REGION Network 1: Header
   // ==============================================================================
   //  Company: Precision Automation & Robotics India Ltd. 
   // ------------------------------------------------------------------------------
   //  Item Code: S21006022015
   //  Author/Created by: Manoj Sonawane
   //  Reviewed/Checked by: Sandip.c
   //  First Release on: 19-07-24
   //  Latest update on:11-03-25
   // ------------------------------------------------------------------------------
   //  Tested with: CPU firmware, model or simulator testing
   //  Engineering/Editor: TIA Portal V17
   // ------------------------------------------------------------------------------
   //  Restrictions:
   //  Dependencies/Requirements:
   //  1. "UDT_IS28xx_To_Plc"
   //  2. "UDT_Plc_To_IS28xx"
   // ------------------------------------------------------------------------------
   //  Change Log:
   //  Ver.	Date		Changed by		Details of changes
   //  1.0	 19-07-24                 Manoj Sonawane            	First release version
   // 1.1              30-09-24                 Harshal Gharmode                         Modify as per shop floor testing
   // 1.2              11-03-25                 Swapnil Asule                                  Remove retry count logic & update                                                                                                                         data Inspection logic
   // ------------------------------------------------------------------------------
   //  Functionality:  : The Cognex In-Sight® 2801 vision system communicates with the Siemence s7-15xx series PLC over Profinet protocol.The main functionality of this block is provided for the user can change the job ID according to their needs and get the inspection result data of Job ID.
   // 
   // 
   //  Inputs
   // iInsightCamera_Input	"UDT_IS28xx_To_Plc"
   // iResetFault	Bool
   // iModuleReset	Bool
   // iAutorunning	Bool
   // iStartJobSelection	Bool
   // iStartInspection	Bool
   // iJobID	Int
   // iUserData	Array[1..60] of Byte
   // iTriggerEnableTimeoutTime	Time
   // iTriggerTimeoutTime	Time
   // iAcquiringTimeOutTime	Time
   // iPrgmNoTimeOut	Time
   // iFeedbackTimeOut	Time
   // 
   //  Outputs
   //  qInsightCamera_Output	"UDT_Plc_To_IS28xx"
   // qJobPass	Bool
   // qJobFail	Bool
   // qJobSelectionOver	Bool
   // qJobInspectionOver	Bool
   // qVisionOnline	Bool
   // qVisionOfflineReason1	Bool
   // qVisionOfflineReason2	Bool
   // qVisionOfflineReason3	Bool
   // qErrBothStartOn	Bool
   // qErrJobSelection	Bool
   // qErrTriggerEnableTimeout	Bool
   // qErrTriggerTimeOut	Bool
   // qErrAcquiringTimeOut	Bool
   // qErrJobIDEchoMismatch	Bool
   // qErrSetUserDataAckNtRcvd	Bool
   // qMsgJobIDMismatch	Bool
   // qInspectionResult	Array[1..60] of Byte
   // 
   //  In-outs
   //  iqRunningJobID	Int
   // ------------------------------------------------------------------------------
   //  Errors reported:
   //  1.qErrTriggerTimeO : Error trigger timeout
   //  2. qErrAcquiringTimeOut;Acquiring Time Out
   //  3. qErrTriggerEnableTimeout:Trigger Enable Time Out
   //  4. qErrJobSelection: Job selection error
   //  5. qErrBothStartOn: Start Inspection & Start Job Selection command are active at same time
   //  6. qErrJobIDEchoMismatch: Set Job ID & its echo is not matched
   //  7. qErrSetUserDataAckNtRcvd: Set user data acknowldge not recived within the defined time.
   // 
   //  Messages reported:
   //   1. qMsgJobIDMismatch: Set Job ID & running JOB ID is not matched
   // ==============================================================================
END_REGION

REGION Network 2: Reset Faults
   // Reset Faults
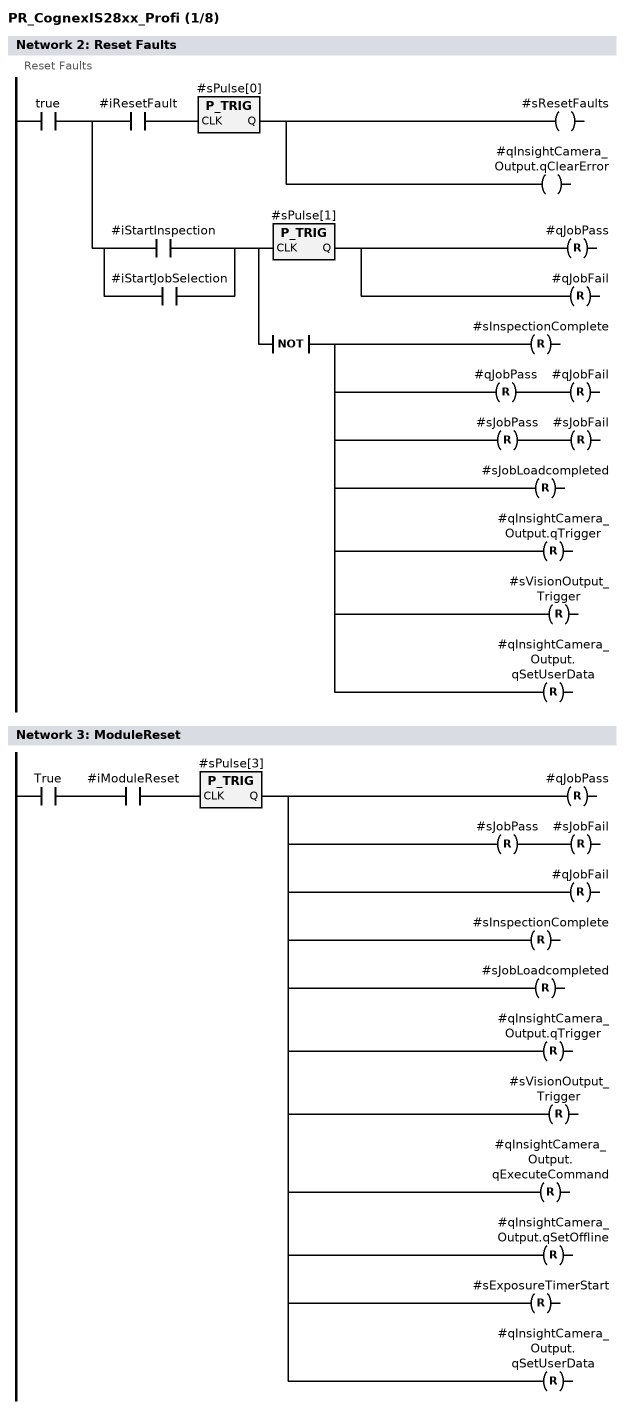
   RUNG wire#powerrail
      Contact( true )
      wire#w1
      Contact( #iResetFault )
      P_Trig( #sPulse[0] )
      wire#w2
      Coil( #sResetFaults )
   END_RUNG
   RUNG wire#w2
      Coil( #qInsightCamera_Output.qClearError )
   END_RUNG
   RUNG wire#w1
      Contact( #iStartInspection )
      wire#w3
      P_Trig( #sPulse[1] )
      wire#w4
      R_Coil( #qJobPass )
   END_RUNG
   RUNG wire#w1
      Contact( #iStartJobSelection )
   END_RUNG wire#w3
   RUNG wire#w4
      R_Coil( #qJobFail )
   END_RUNG
   RUNG wire#w3
      Not()
      wire#w5
      R_Coil( #sInspectionComplete )
   END_RUNG
   RUNG wire#w5
      R_Coil( #qJobPass )
      R_Coil( #qJobFail )
   END_RUNG
   RUNG wire#w5
      R_Coil( #sJobPass )
      R_Coil( #sJobFail )
   END_RUNG
   RUNG wire#w5
      R_Coil( #sJobLoadcompleted )
   END_RUNG
   RUNG wire#w5
      R_Coil( #qInsightCamera_Output.qTrigger )
   END_RUNG
   RUNG wire#w5
      R_Coil( #sVisionOutput_Trigger )
   END_RUNG
   RUNG wire#w5
      R_Coil( #qInsightCamera_Output.qSetUserData )
   END_RUNG
   // the same network as SCL:
   #_w1 := true AND #iResetFault;
   #_w2 := #_w1 AND NOT #sPulse[0];   // rising edge
   #sPulse[0] := #_w1;
   #sResetFaults := #_w2;
   #qInsightCamera_Output.qClearError := #_w2;
   #_w3 := true AND (#iStartInspection OR #iStartJobSelection);
   #_w4 := #_w3 AND NOT #sPulse[1];   // rising edge
   #sPulse[1] := #_w3;
   IF #_w4 THEN
       #qJobPass := FALSE;
       #qJobFail := FALSE;
   END_IF;
   IF NOT #_w3 THEN
       #sInspectionComplete := FALSE;
       #qJobPass := FALSE;
       #qJobFail := FALSE;
       #sJobPass := FALSE;
       #sJobFail := FALSE;
       #sJobLoadcompleted := FALSE;
       #qInsightCamera_Output.qTrigger := FALSE;
       #sVisionOutput_Trigger := FALSE;
       #qInsightCamera_Output.qSetUserData := FALSE;
   END_IF;
END_REGION

REGION Network 3: ModuleReset
   RUNG wire#powerrail
      Contact( True )
      Contact( #iModuleReset )
      P_Trig( #sPulse[3] )
      wire#w1
      R_Coil( #qJobPass )
   END_RUNG
   RUNG wire#w1
      R_Coil( #sJobPass )
      R_Coil( #sJobFail )
   END_RUNG
   RUNG wire#w1
      R_Coil( #qJobFail )
   END_RUNG
   RUNG wire#w1
      R_Coil( #sInspectionComplete )
   END_RUNG
   RUNG wire#w1
      R_Coil( #sJobLoadcompleted )
   END_RUNG
   RUNG wire#w1
      R_Coil( #qInsightCamera_Output.qTrigger )
   END_RUNG
   RUNG wire#w1
      R_Coil( #sVisionOutput_Trigger )
   END_RUNG
   RUNG wire#w1
      R_Coil( #qInsightCamera_Output.qExecuteCommand )
   END_RUNG
   RUNG wire#w1
      R_Coil( #qInsightCamera_Output.qSetOffline )
   END_RUNG
   RUNG wire#w1
      R_Coil( #sExposureTimerStart )
   END_RUNG
   RUNG wire#w1
      R_Coil( #qInsightCamera_Output.qSetUserData )
   END_RUNG
   // the same network as SCL:
   #_w1 := True AND #iModuleReset;
   #_w2 := #_w1 AND NOT #sPulse[3];   // rising edge
   #sPulse[3] := #_w1;
   IF #_w2 THEN
       #qJobPass := FALSE;
       #sJobPass := FALSE;
       #sJobFail := FALSE;
       #qJobFail := FALSE;
       #sInspectionComplete := FALSE;
       #sJobLoadcompleted := FALSE;
       #qInsightCamera_Output.qTrigger := FALSE;
       #sVisionOutput_Trigger := FALSE;
       #qInsightCamera_Output.qExecuteCommand := FALSE;
       #qInsightCamera_Output.qSetOffline := FALSE;
       #sExposureTimerStart := FALSE;
       #qInsightCamera_Output.qSetUserData := FALSE;
   END_IF;
END_REGION

REGION Network 4: Time out validation
   // Time out validation 1. Trigger enable time out
   // 2. Trigger time out
   // 3. Acquiring TimeOut Time
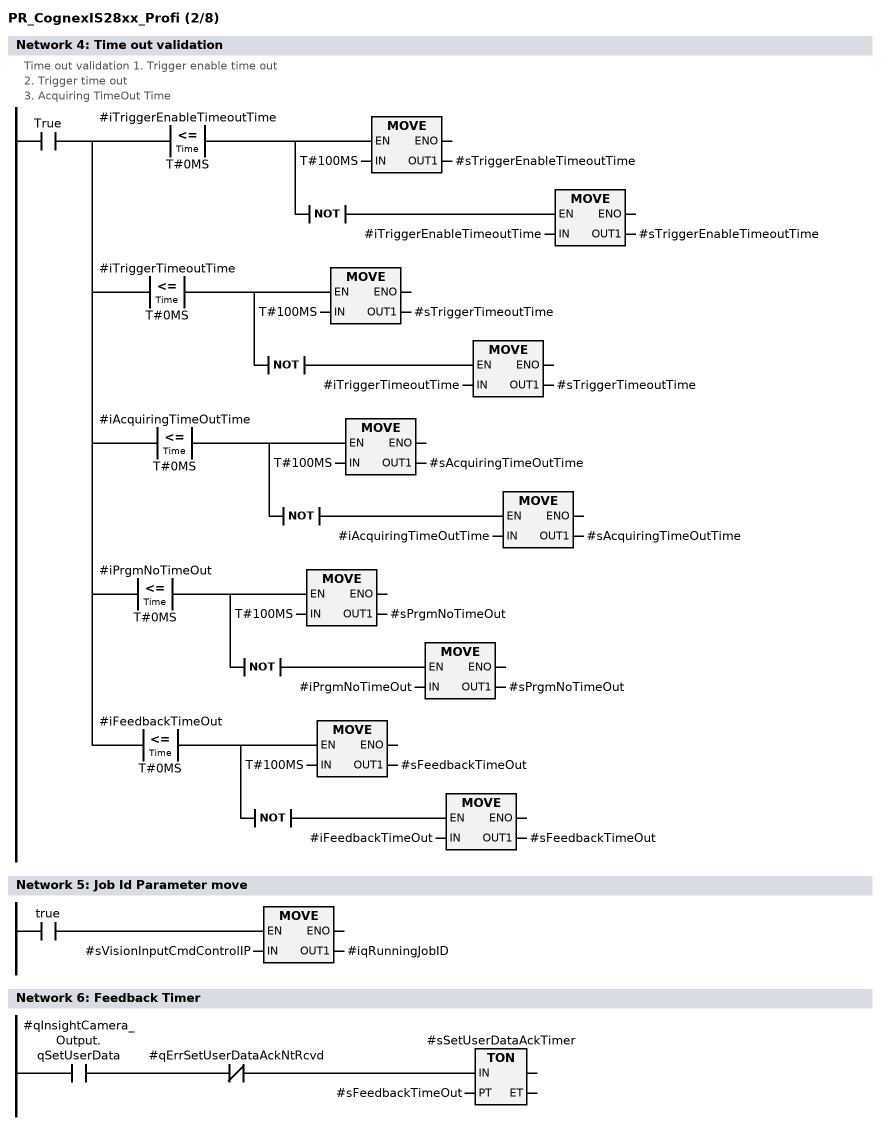
   RUNG wire#powerrail
      Contact( True )
      wire#w1
      { S7_Templates := "SrcType := Time" } LE_Contact(in1 := #iTriggerEnableTimeoutTime, in2 := T#0MS)
      wire#w2
      Move(in := T#100MS, out1 => #sTriggerEnableTimeoutTime)
   END_RUNG
   RUNG wire#w2
      Not()
      Move(in := #iTriggerEnableTimeoutTime, out1 => #sTriggerEnableTimeoutTime)
   END_RUNG
   RUNG wire#w1
      { S7_Templates := "SrcType := Time" } LE_Contact(in1 := #iTriggerTimeoutTime, in2 := T#0MS)
      wire#w3
      Move(in := T#100MS, out1 => #sTriggerTimeoutTime)
   END_RUNG
   RUNG wire#w3
      Not()
      Move(in := #iTriggerTimeoutTime, out1 => #sTriggerTimeoutTime)
   END_RUNG
   RUNG wire#w1
      { S7_Templates := "SrcType := Time" } LE_Contact(in1 := #iAcquiringTimeOutTime, in2 := T#0MS)
      wire#w4
      Move(in := T#100MS, out1 => #sAcquiringTimeOutTime)
   END_RUNG
   RUNG wire#w4
      Not()
      Move(in := #iAcquiringTimeOutTime, out1 => #sAcquiringTimeOutTime)
   END_RUNG
   RUNG wire#w1
      { S7_Templates := "SrcType := Time" } LE_Contact(in1 := #iPrgmNoTimeOut, in2 := T#0MS)
      wire#w5
      Move(in := T#100MS, out1 => #sPrgmNoTimeOut)
   END_RUNG
   RUNG wire#w5
      Not()
      Move(in := #iPrgmNoTimeOut, out1 => #sPrgmNoTimeOut)
   END_RUNG
   RUNG wire#w1
      { S7_Templates := "SrcType := Time" } LE_Contact(in1 := #iFeedbackTimeOut, in2 := T#0MS)
      wire#w6
      Move(in := T#100MS, out1 => #sFeedbackTimeOut)
   END_RUNG
   RUNG wire#w6
      Not()
      Move(in := #iFeedbackTimeOut, out1 => #sFeedbackTimeOut)
   END_RUNG
   // the same network as SCL:
   #_w1 := True AND (#iTriggerEnableTimeoutTime <= T#0MS);
   IF #_w1 THEN #sTriggerEnableTimeoutTime := T#100MS; END_IF;
   IF NOT #_w1 THEN #sTriggerEnableTimeoutTime := #iTriggerEnableTimeoutTime; END_IF;
   #_w2 := True AND (#iTriggerTimeoutTime <= T#0MS);
   IF #_w2 THEN #sTriggerTimeoutTime := T#100MS; END_IF;
   IF NOT #_w2 THEN #sTriggerTimeoutTime := #iTriggerTimeoutTime; END_IF;
   #_w3 := True AND (#iAcquiringTimeOutTime <= T#0MS);
   IF #_w3 THEN #sAcquiringTimeOutTime := T#100MS; END_IF;
   IF NOT #_w3 THEN #sAcquiringTimeOutTime := #iAcquiringTimeOutTime; END_IF;
   #_w4 := True AND (#iPrgmNoTimeOut <= T#0MS);
   IF #_w4 THEN #sPrgmNoTimeOut := T#100MS; END_IF;
   IF NOT #_w4 THEN #sPrgmNoTimeOut := #iPrgmNoTimeOut; END_IF;
   #_w5 := True AND (#iFeedbackTimeOut <= T#0MS);
   IF #_w5 THEN #sFeedbackTimeOut := T#100MS; END_IF;
   IF NOT #_w5 THEN #sFeedbackTimeOut := #iFeedbackTimeOut; END_IF;
END_REGION

REGION Network 5: Job Id Parameter move
   RUNG wire#powerrail
      Contact( true )
      Move(in := #sVisionInputCmdControlIP, out1 => #iqRunningJobID)
   END_RUNG
   // the same network as SCL:
   IF true THEN #iqRunningJobID := #sVisionInputCmdControlIP; END_IF;
END_REGION

REGION Network 6: Feedback Timer
   #sSetUserDataAckTimer(IN := #qInsightCamera_Output.qSetUserData AND NOT #qErrSetUserDataAckNtRcvd,   // TON
                         PT := #sFeedbackTimeOut);
END_REGION

REGION Network 7: UserData
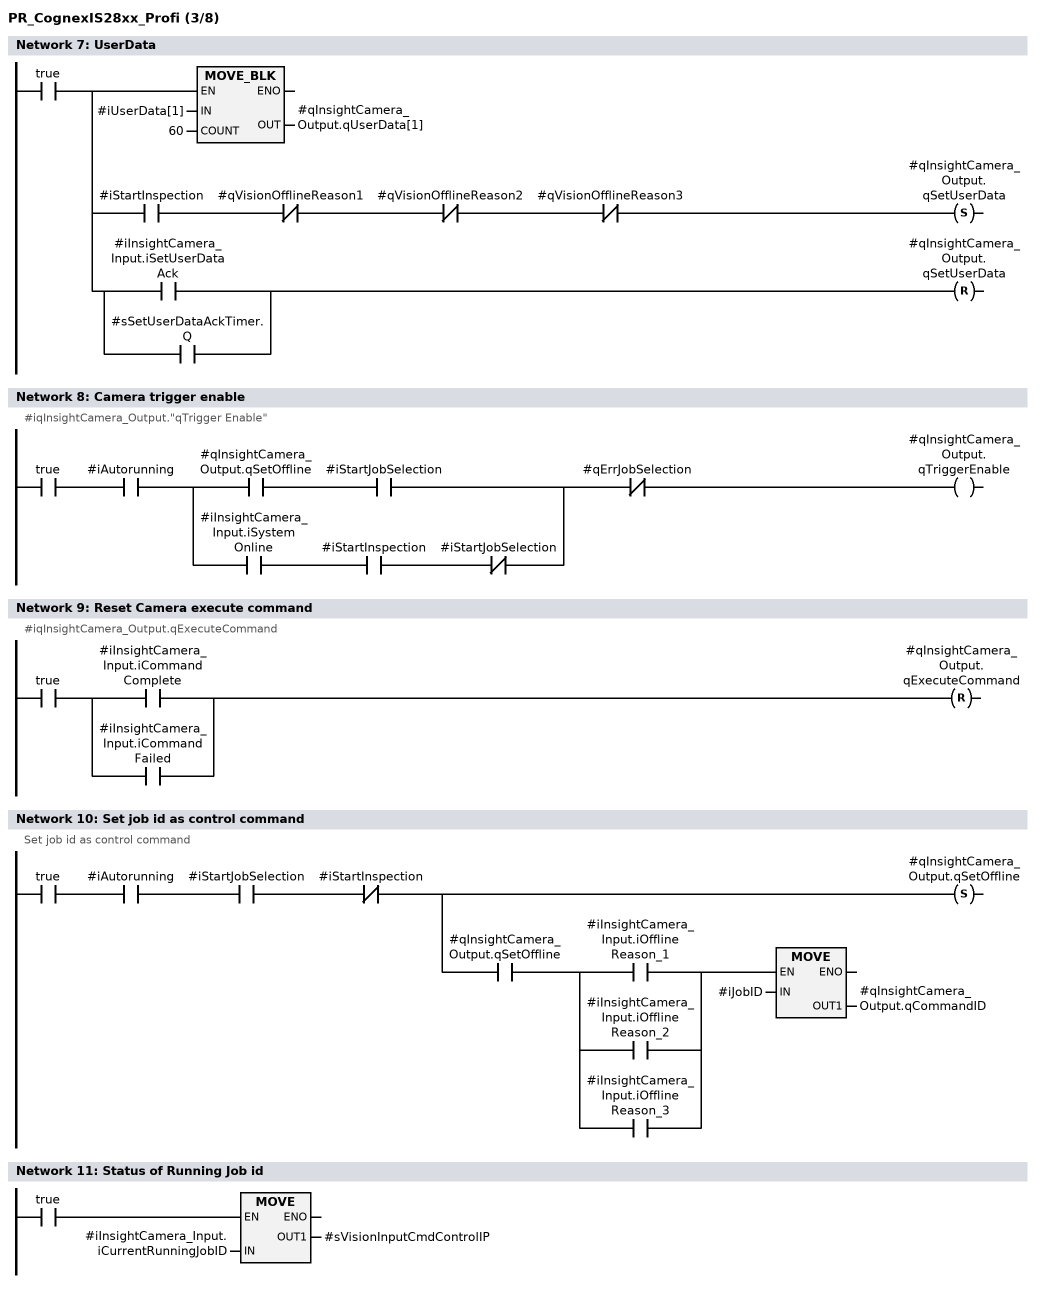
   IF true THEN
       MOVE_BLK(IN := #iUserData[1], COUNT := 60, OUT => #qInsightCamera_Output.qUserData[1]);
   END_IF;
   IF true AND #iStartInspection AND NOT #qVisionOfflineReason1 AND NOT #qVisionOfflineReason2 AND NOT #qVisionOfflineReason3 THEN
       #qInsightCamera_Output.qSetUserData := TRUE;
   END_IF;
   IF true AND (#iInsightCamera_Input.iSetUserDataAck OR #sSetUserDataAckTimer.Q) THEN
       #qInsightCamera_Output.qSetUserData := FALSE;
   END_IF;
END_REGION

REGION Network 8: Camera trigger enable
   // #iqInsightCamera_Output."qTrigger Enable"
   RUNG wire#powerrail
      Contact( true )
      Contact( #iAutorunning )
      wire#w1
      Contact( #qInsightCamera_Output.qSetOffline )
      Contact( #iStartJobSelection )
      wire#w2
      I_Contact( #qErrJobSelection )
      Coil( #qInsightCamera_Output.qTriggerEnable )
   END_RUNG
   RUNG wire#w1
      Contact( #iInsightCamera_Input.iSystemOnline )
      Contact( #iStartInspection )
      I_Contact( #iStartJobSelection )
   END_RUNG wire#w2
   // the same network as SCL:
   #qInsightCamera_Output.qTriggerEnable := true AND #iAutorunning AND ((#qInsightCamera_Output.qSetOffline AND #iStartJobSelection) OR (#iInsightCamera_Input.iSystemOnline AND #iStartInspection AND NOT #iStartJobSelection)) AND NOT #qErrJobSelection;
END_REGION

REGION Network 9: Reset Camera execute command
   // #iqInsightCamera_Output.qExecuteCommand
   RUNG wire#powerrail
      Contact( true )
      wire#w1
      Contact( #iInsightCamera_Input.iCommandComplete )
      wire#w2
      R_Coil( #qInsightCamera_Output.qExecuteCommand )
   END_RUNG
   RUNG wire#w1
      Contact( #iInsightCamera_Input.iCommandFailed )
   END_RUNG wire#w2
   // the same network as SCL:
   IF true AND (#iInsightCamera_Input.iCommandComplete OR #iInsightCamera_Input.iCommandFailed) THEN
       #qInsightCamera_Output.qExecuteCommand := FALSE;
   END_IF;
END_REGION

REGION Network 10: Set job id as control command
   // Set job id as control command
   RUNG wire#powerrail
      Contact( true )
      Contact( #iAutorunning )
      Contact( #iStartJobSelection )
      I_Contact( #iStartInspection )
      wire#w1
      S_Coil( #qInsightCamera_Output.qSetOffline )
   END_RUNG
   RUNG wire#w1
      Contact( #qInsightCamera_Output.qSetOffline )
      wire#w2
      Contact( #iInsightCamera_Input.iOfflineReason_1 )
      wire#w3
      Move(in := #iJobID, out1 => #qInsightCamera_Output.qCommandID)
   END_RUNG
   RUNG wire#w2
      Contact( #iInsightCamera_Input.iOfflineReason_2 )
   END_RUNG wire#w3
   RUNG wire#w2
      Contact( #iInsightCamera_Input.iOfflineReason_3 )
   END_RUNG wire#w3
   // the same network as SCL:
   #_w1 := true AND #iAutorunning AND #iStartJobSelection AND NOT #iStartInspection;
   IF #_w1 THEN #qInsightCamera_Output.qSetOffline := TRUE; END_IF;
   IF #_w1 AND #qInsightCamera_Output.qSetOffline AND (#iInsightCamera_Input.iOfflineReason_1 OR #iInsightCamera_Input.iOfflineReason_2 OR #iInsightCamera_Input.iOfflineReason_3) THEN
       #qInsightCamera_Output.qCommandID := #iJobID;
   END_IF;
END_REGION

REGION Network 11: Status of Running Job id
   RUNG wire#powerrail
      Contact( true )
      Move(in := #iInsightCamera_Input.iCurrentRunningJobID, out1 => #sVisionInputCmdControlIP)
   END_RUNG
   // the same network as SCL:
   IF true THEN #sVisionInputCmdControlIP := #iInsightCamera_Input.iCurrentRunningJobID; END_IF;
END_REGION

REGION Network 12: Set Execute command as per Job selection
   // Set Execute command as per Job selection
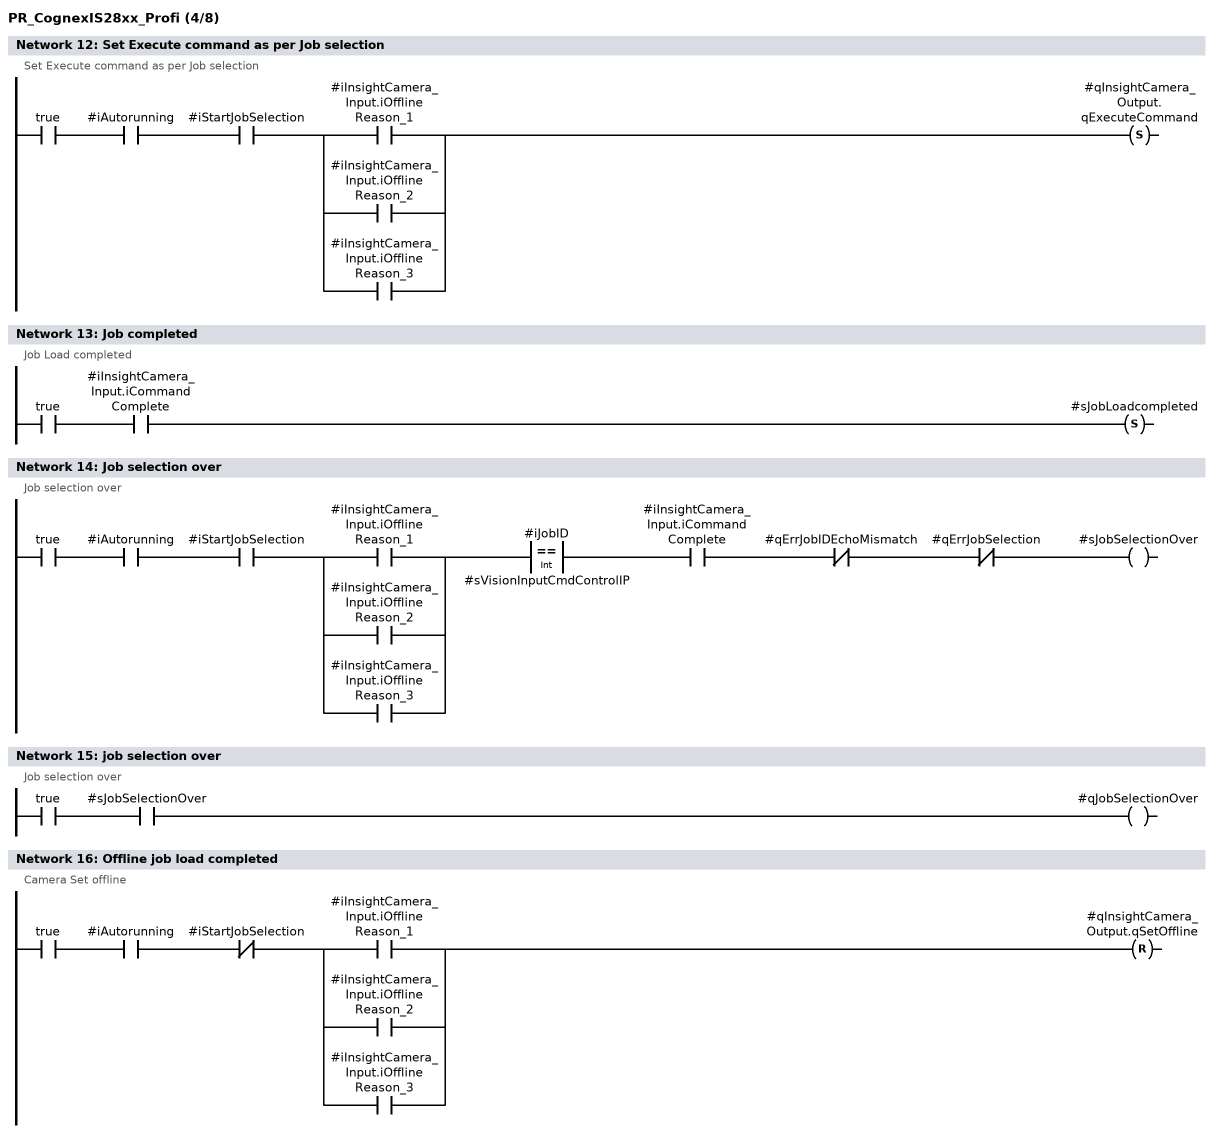
   RUNG wire#powerrail
      Contact( true )
      Contact( #iAutorunning )
      Contact( #iStartJobSelection )
      wire#w1
      Contact( #iInsightCamera_Input.iOfflineReason_1 )
      wire#w2
      S_Coil( #qInsightCamera_Output.qExecuteCommand )
   END_RUNG
   RUNG wire#w1
      Contact( #iInsightCamera_Input.iOfflineReason_2 )
   END_RUNG wire#w2
   RUNG wire#w1
      Contact( #iInsightCamera_Input.iOfflineReason_3 )
   END_RUNG wire#w2
   // the same network as SCL:
   IF true AND #iAutorunning AND #iStartJobSelection AND (#iInsightCamera_Input.iOfflineReason_1 OR #iInsightCamera_Input.iOfflineReason_2 OR #iInsightCamera_Input.iOfflineReason_3) THEN
       #qInsightCamera_Output.qExecuteCommand := TRUE;
   END_IF;
END_REGION

REGION Network 13: Job completed
   // Job Load completed
   RUNG wire#powerrail
      Contact( true )
      Contact( #iInsightCamera_Input.iCommandComplete )
      S_Coil( #sJobLoadcompleted )
   END_RUNG
   // the same network as SCL:
   IF true AND #iInsightCamera_Input.iCommandComplete THEN #sJobLoadcompleted := TRUE; END_IF;
END_REGION

REGION Network 14: Job selection over
   // Job selection over
   RUNG wire#powerrail
      Contact( true )
      Contact( #iAutorunning )
      Contact( #iStartJobSelection )
      wire#w1
      Contact( #iInsightCamera_Input.iOfflineReason_1 )
      wire#w2
      { S7_Templates := "SrcType := Int" } EQ_Contact(in1 := #iJobID, in2 := #sVisionInputCmdControlIP)
      Contact( #iInsightCamera_Input.iCommandComplete )
      I_Contact( #qErrJobIDEchoMismatch )
      I_Contact( #qErrJobSelection )
      Coil( #sJobSelectionOver )
   END_RUNG
   RUNG wire#w1
      Contact( #iInsightCamera_Input.iOfflineReason_2 )
   END_RUNG wire#w2
   RUNG wire#w1
      Contact( #iInsightCamera_Input.iOfflineReason_3 )
   END_RUNG wire#w2
   // the same network as SCL:
   #sJobSelectionOver := true AND #iAutorunning AND #iStartJobSelection AND (#iInsightCamera_Input.iOfflineReason_1 OR #iInsightCamera_Input.iOfflineReason_2 OR #iInsightCamera_Input.iOfflineReason_3) AND (#iJobID = #sVisionInputCmdControlIP) AND #iInsightCamera_Input.iCommandComplete AND NOT #qErrJobIDEchoMismatch AND NOT #qErrJobSelection;
END_REGION

REGION Network 15: job selection over
   // Job selection over
   RUNG wire#powerrail
      Contact( true )
      Contact( #sJobSelectionOver )
      Coil( #qJobSelectionOver )
   END_RUNG
   // the same network as SCL:
   #qJobSelectionOver := true AND #sJobSelectionOver;
END_REGION

REGION Network 16: Offline job load completed
   // Camera Set offline
   RUNG wire#powerrail
      Contact( true )
      Contact( #iAutorunning )
      I_Contact( #iStartJobSelection )
      wire#w1
      Contact( #iInsightCamera_Input.iOfflineReason_1 )
      wire#w2
      R_Coil( #qInsightCamera_Output.qSetOffline )
   END_RUNG
   RUNG wire#w1
      Contact( #iInsightCamera_Input.iOfflineReason_2 )
   END_RUNG wire#w2
   RUNG wire#w1
      Contact( #iInsightCamera_Input.iOfflineReason_3 )
   END_RUNG wire#w2
   // the same network as SCL:
   IF true AND #iAutorunning AND NOT #iStartJobSelection AND (#iInsightCamera_Input.iOfflineReason_1 OR #iInsightCamera_Input.iOfflineReason_2 OR #iInsightCamera_Input.iOfflineReason_3) THEN
       #qInsightCamera_Output.qSetOffline := FALSE;
   END_IF;
END_REGION

REGION Network 17: Trigger Enable
   // Trigger Enable
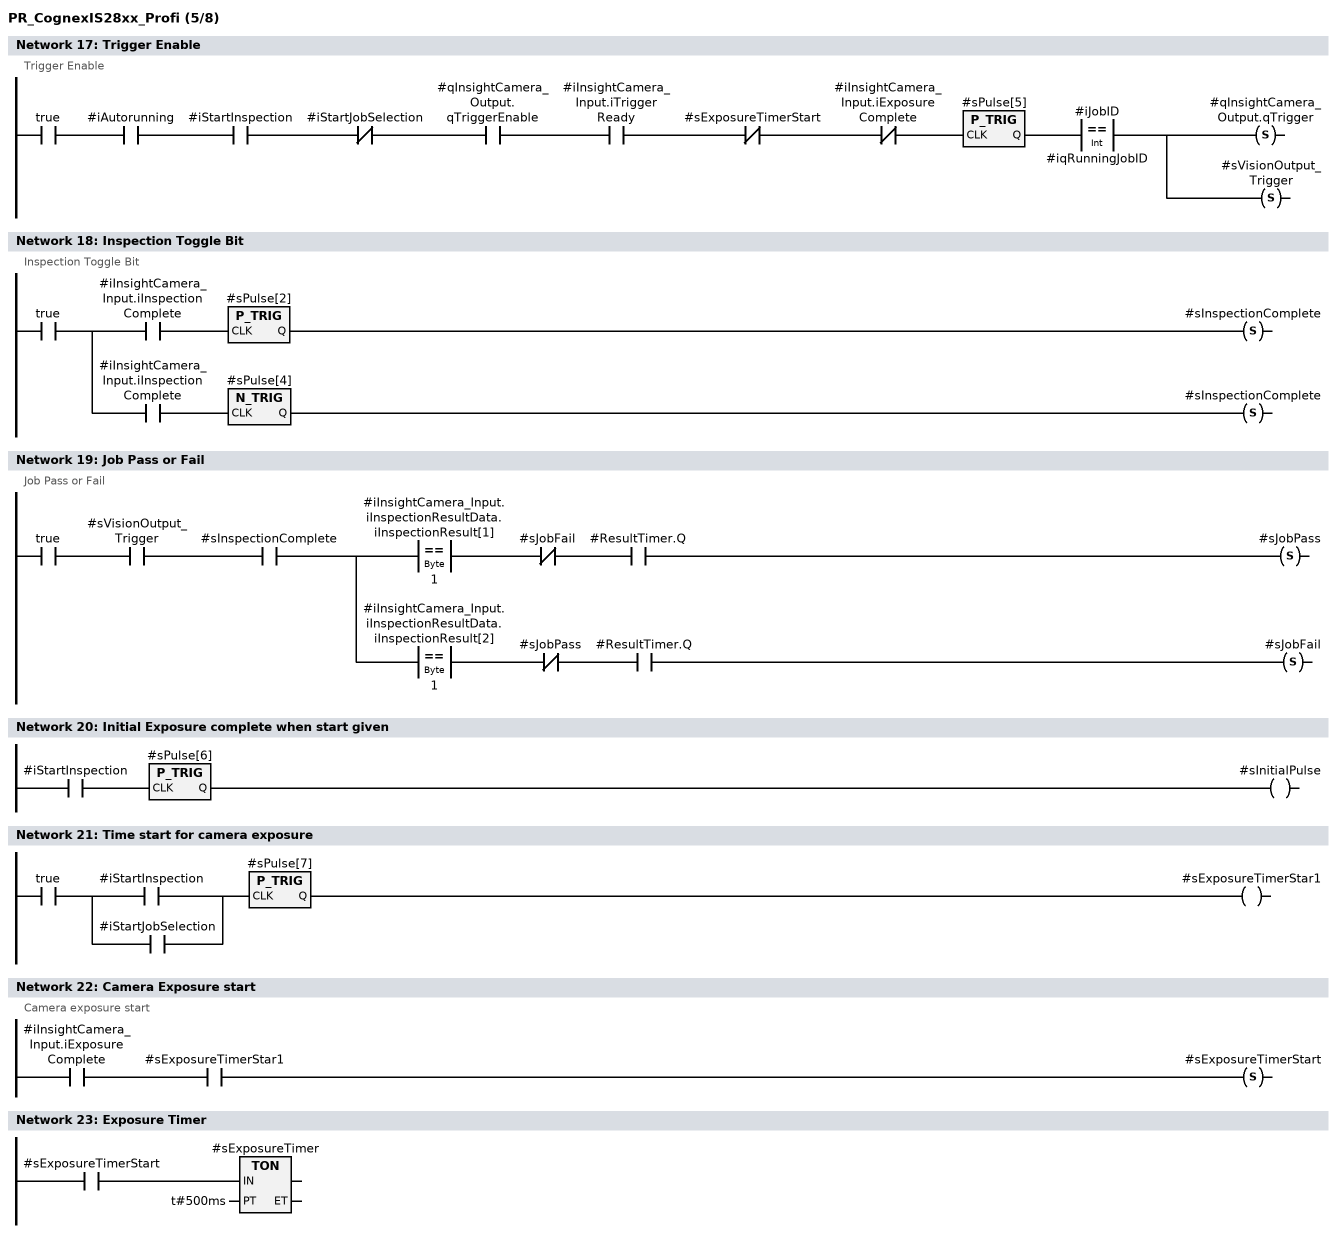
   RUNG wire#powerrail
      Contact( true )
      Contact( #iAutorunning )
      Contact( #iStartInspection )
      I_Contact( #iStartJobSelection )
      Contact( #qInsightCamera_Output.qTriggerEnable )
      Contact( #iInsightCamera_Input.iTriggerReady )
      I_Contact( #sExposureTimerStart )
      I_Contact( #iInsightCamera_Input.iExposureComplete )
      P_Trig( #sPulse[5] )
      { S7_Templates := "SrcType := Int" } EQ_Contact(in1 := #iJobID, in2 := #iqRunningJobID)
      wire#w1
      S_Coil( #qInsightCamera_Output.qTrigger )
   END_RUNG
   RUNG wire#w1
      S_Coil( #sVisionOutput_Trigger )
   END_RUNG
   // the same network as SCL:
   #_w1 := true AND #iAutorunning AND #iStartInspection AND NOT #iStartJobSelection AND #qInsightCamera_Output.qTriggerEnable AND #iInsightCamera_Input.iTriggerReady AND NOT #sExposureTimerStart AND NOT #iInsightCamera_Input.iExposureComplete;
   #_w2 := #_w1 AND NOT #sPulse[5];   // rising edge
   #sPulse[5] := #_w1;
   IF #_w2 AND (#iJobID = #iqRunningJobID) THEN
       #qInsightCamera_Output.qTrigger := TRUE;
       #sVisionOutput_Trigger := TRUE;
   END_IF;
END_REGION

REGION Network 18: Inspection Toggle Bit
   // Inspection Toggle Bit
   RUNG wire#powerrail
      Contact( true )
      wire#w1
      Contact( #iInsightCamera_Input.iInspectionComplete )
      P_Trig( #sPulse[2] )
      S_Coil( #sInspectionComplete )
   END_RUNG
   RUNG wire#w1
      Contact( #iInsightCamera_Input.iInspectionComplete )
      N_Trig( #sPulse[4] )
      S_Coil( #sInspectionComplete )
   END_RUNG
   // the same network as SCL:
   #_w1 := true AND #iInsightCamera_Input.iInspectionComplete;
   #_w2 := #_w1 AND NOT #sPulse[2];   // rising edge
   #sPulse[2] := #_w1;
   IF #_w2 THEN #sInspectionComplete := TRUE; END_IF;
   #_w3 := true AND #iInsightCamera_Input.iInspectionComplete;
   #_w4 := NOT #_w3 AND #sPulse[4];   // falling edge
   #sPulse[4] := #_w3;
   IF #_w4 THEN #sInspectionComplete := TRUE; END_IF;
END_REGION

REGION Network 19: Job Pass or Fail
   // Job Pass or Fail
   RUNG wire#powerrail
      Contact( true )
      Contact( #sVisionOutput_Trigger )
      Contact( #sInspectionComplete )
      wire#w1
      { S7_Templates := "SrcType := Byte" } EQ_Contact(in1 := #iInsightCamera_Input.iInspectionResultData.iInspectionResult[1], in2 := 1)
      I_Contact( #sJobFail )
      Contact( #ResultTimer.Q )
      S_Coil( #sJobPass )
   END_RUNG
   RUNG wire#w1
      { S7_Templates := "SrcType := Byte" } EQ_Contact(in1 := #iInsightCamera_Input.iInspectionResultData.iInspectionResult[2], in2 := 1)
      I_Contact( #sJobPass )
      Contact( #ResultTimer.Q )
      S_Coil( #sJobFail )
   END_RUNG
   // the same network as SCL:
   #_w1 := true AND #sVisionOutput_Trigger AND #sInspectionComplete;
   IF #_w1 AND (#iInsightCamera_Input.iInspectionResultData.iInspectionResult[1] = 1) AND NOT #sJobFail AND #ResultTimer.Q THEN
       #sJobPass := TRUE;
   END_IF;
   IF #_w1 AND (#iInsightCamera_Input.iInspectionResultData.iInspectionResult[2] = 1) AND NOT #sJobPass AND #ResultTimer.Q THEN
       #sJobFail := TRUE;
   END_IF;
END_REGION

REGION Network 20: Initial Exposure complete when start given
   RUNG wire#powerrail
      Contact( #iStartInspection )
      P_Trig( #sPulse[6] )
      Coil( #sInitialPulse )
   END_RUNG
   // the same network as SCL:
   #_w1 := #iStartInspection AND NOT #sPulse[6];   // rising edge
   #sPulse[6] := #iStartInspection;
   #sInitialPulse := #_w1;
END_REGION

REGION Network 21: Time start for camera exposure
   RUNG wire#powerrail
      Contact( true )
      wire#w1
      Contact( #iStartInspection )
      wire#w2
      P_Trig( #sPulse[7] )
      Coil( #sExposureTimerStar1 )
   END_RUNG
   RUNG wire#w1
      Contact( #iStartJobSelection )
   END_RUNG wire#w2
   // the same network as SCL:
   #_w1 := true AND (#iStartInspection OR #iStartJobSelection);
   #_w2 := #_w1 AND NOT #sPulse[7];   // rising edge
   #sPulse[7] := #_w1;
   #sExposureTimerStar1 := #_w2;
END_REGION

REGION Network 22: Camera Exposure start
   // Camera exposure start
   RUNG wire#powerrail
      Contact( #iInsightCamera_Input.iExposureComplete )
      Contact( #sExposureTimerStar1 )
      S_Coil( #sExposureTimerStart )
   END_RUNG
   // the same network as SCL:
   IF #iInsightCamera_Input.iExposureComplete AND #sExposureTimerStar1 THEN
       #sExposureTimerStart := TRUE;
   END_IF;
END_REGION

REGION Network 23: Exposure Timer
   #sExposureTimer(IN := #sExposureTimerStart, PT := t#500ms);   // TON
END_REGION

REGION Network 24: Exposure Timer Complete
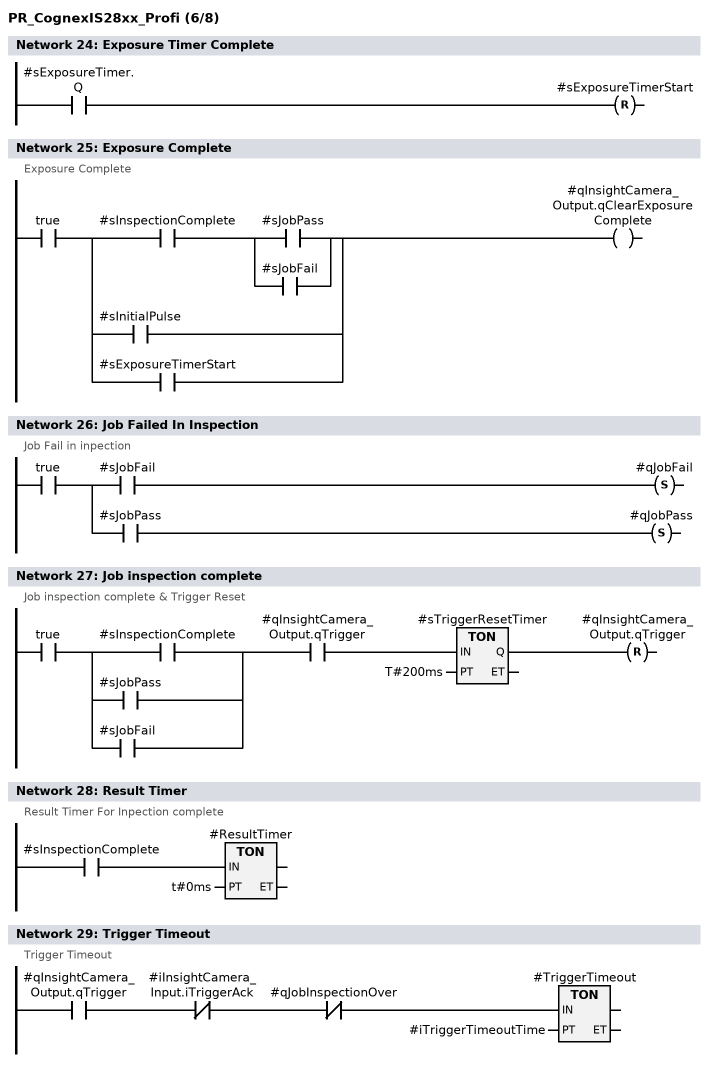
   RUNG wire#powerrail
      Contact( #sExposureTimer.Q )
      R_Coil( #sExposureTimerStart )
   END_RUNG
   // the same network as SCL:
   IF #sExposureTimer.Q THEN #sExposureTimerStart := FALSE; END_IF;
END_REGION

REGION Network 25: Exposure Complete
   // Exposure Complete
   RUNG wire#powerrail
      Contact( true )
      wire#w1
      Contact( #sInspectionComplete )
      wire#w2
      Contact( #sJobPass )
      wire#w3
      Coil( #qInsightCamera_Output.qClearExposureComplete )
   END_RUNG
   RUNG wire#w2
      Contact( #sJobFail )
   END_RUNG wire#w3
   RUNG wire#w1
      Contact( #sInitialPulse )
   END_RUNG wire#w3
   RUNG wire#w1
      Contact( #sExposureTimerStart )
   END_RUNG wire#w3
   // the same network as SCL:
   #qInsightCamera_Output.qClearExposureComplete := true AND ((#sInspectionComplete AND (#sJobPass OR #sJobFail)) OR #sInitialPulse OR #sExposureTimerStart);
END_REGION

REGION Network 26: Job Failed In Inspection
   // Job Fail in inpection
   RUNG wire#powerrail
      Contact( true )
      wire#w1
      Contact( #sJobFail )
      S_Coil( #qJobFail )
   END_RUNG
   RUNG wire#w1
      Contact( #sJobPass )
      S_Coil( #qJobPass )
   END_RUNG
   // the same network as SCL:
   IF true AND #sJobFail THEN #qJobFail := TRUE; END_IF;
   IF true AND #sJobPass THEN #qJobPass := TRUE; END_IF;
END_REGION

REGION Network 27: Job inspection complete
   // Job inspection complete & Trigger Reset
   #sTriggerResetTimer(IN := true AND (#sInspectionComplete OR #sJobPass OR #sJobFail) AND #qInsightCamera_Output.qTrigger,   // TON
                       PT := T#200ms);
   IF #sTriggerResetTimer.Q THEN #qInsightCamera_Output.qTrigger := FALSE; END_IF;
END_REGION

REGION Network 28: Result Timer
   // Result Timer For Inpection complete
   #ResultTimer(IN := #sInspectionComplete, PT := t#0ms);   // TON
END_REGION

REGION Network 29: Trigger Timeout
   // Trigger Timeout
   #TriggerTimeout(IN := #qInsightCamera_Output.qTrigger AND NOT #iInsightCamera_Input.iTriggerAck AND NOT #qJobInspectionOver,   // TON
                   PT := #iTriggerTimeoutTime);
END_REGION

REGION Network 30: Trigger Enable TimeOut
   // Trigger Enable TimeOut
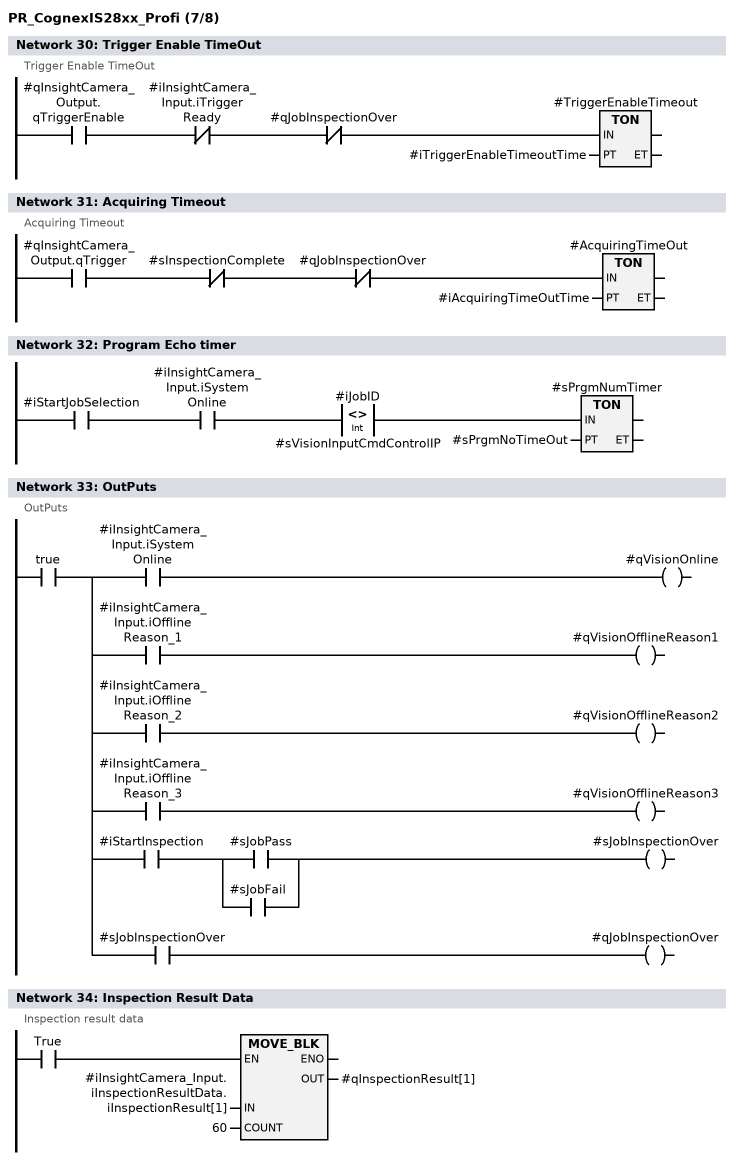
   #TriggerEnableTimeout(IN := #qInsightCamera_Output.qTriggerEnable AND NOT #iInsightCamera_Input.iTriggerReady AND NOT #qJobInspectionOver,   // TON
                         PT := #iTriggerEnableTimeoutTime);
END_REGION

REGION Network 31: Acquiring Timeout
   // Acquiring Timeout
   #AcquiringTimeOut(IN := #qInsightCamera_Output.qTrigger AND NOT #sInspectionComplete AND NOT #qJobInspectionOver,   // TON
                     PT := #iAcquiringTimeOutTime);
END_REGION

REGION Network 32: Program Echo timer
   #sPrgmNumTimer(IN := #iStartJobSelection AND #iInsightCamera_Input.iSystemOnline AND (#iJobID <> #sVisionInputCmdControlIP),   // TON
                  PT := #sPrgmNoTimeOut);
END_REGION

REGION Network 33: OutPuts
   // OutPuts
   RUNG wire#powerrail
      Contact( true )
      wire#w1
      Contact( #iInsightCamera_Input.iSystemOnline )
      Coil( #qVisionOnline )
   END_RUNG
   RUNG wire#w1
      Contact( #iInsightCamera_Input.iOfflineReason_1 )
      Coil( #qVisionOfflineReason1 )
   END_RUNG
   RUNG wire#w1
      Contact( #iInsightCamera_Input.iOfflineReason_2 )
      Coil( #qVisionOfflineReason2 )
   END_RUNG
   RUNG wire#w1
      Contact( #iInsightCamera_Input.iOfflineReason_3 )
      Coil( #qVisionOfflineReason3 )
   END_RUNG
   RUNG wire#w1
      Contact( #iStartInspection )
      wire#w2
      Contact( #sJobPass )
      wire#w3
      Coil( #sJobInspectionOver )
   END_RUNG
   RUNG wire#w2
      Contact( #sJobFail )
   END_RUNG wire#w3
   RUNG wire#w1
      Contact( #sJobInspectionOver )
      Coil( #qJobInspectionOver )
   END_RUNG
   // the same network as SCL:
   #qVisionOnline := true AND #iInsightCamera_Input.iSystemOnline;
   #qVisionOfflineReason1 := true AND #iInsightCamera_Input.iOfflineReason_1;
   #qVisionOfflineReason2 := true AND #iInsightCamera_Input.iOfflineReason_2;
   #qVisionOfflineReason3 := true AND #iInsightCamera_Input.iOfflineReason_3;
   #sJobInspectionOver := true AND #iStartInspection AND (#sJobPass OR #sJobFail);
   #qJobInspectionOver := true AND #sJobInspectionOver;
END_REGION

REGION Network 34: Inspection Result Data
   // Inspection result data
   IF True THEN
       MOVE_BLK(IN := #iInsightCamera_Input.iInspectionResultData.iInspectionResult[1],
                COUNT := 60,
                OUT => #qInspectionResult[1]);
   END_IF;
END_REGION

REGION Network 35: Errors
   // Errors: 
   // qErrTriggerTimeOut: Tigger TimeOut Error Occured
   // qErrAcquiringTimeout: Acquiring TimeOut Error Occured
   // qErrTriggerEnableTimeout: Trigger Enable TimeOut Occured
   // #qErrJobIDEchoMismatch:Job ID Echo Mismatch
   // #qErrJobSelection: Job Error Selection wrong
   // #qErrBothStartOn:Job selection and job inspection both command at time
   // #qErrRetryCount: Retry count value Not set
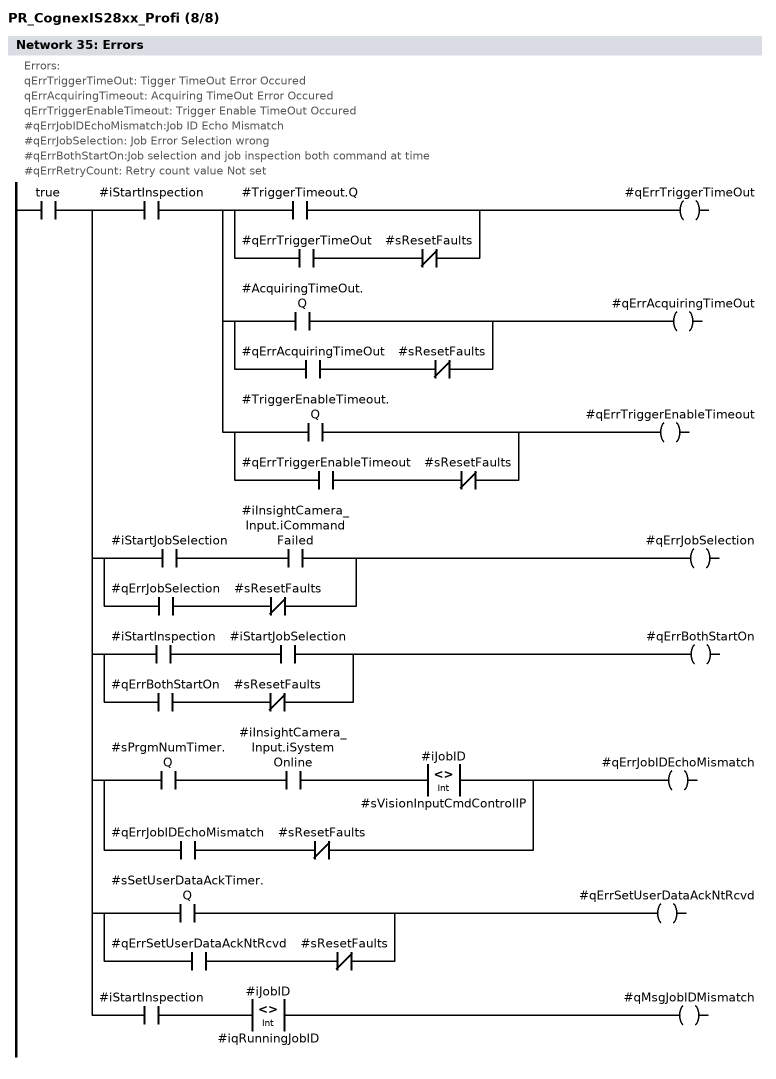
   RUNG wire#powerrail
      Contact( true )
      wire#w1
      Contact( #iStartInspection )
      wire#w2
      Contact( #TriggerTimeout.Q )
      wire#w3
      Coil( #qErrTriggerTimeOut )
   END_RUNG
   RUNG wire#w2
      Contact( #qErrTriggerTimeOut )
      I_Contact( #sResetFaults )
   END_RUNG wire#w3
   RUNG wire#w2
      Contact( #AcquiringTimeOut.Q )
      wire#w4
      Coil( #qErrAcquiringTimeOut )
   END_RUNG
   RUNG wire#w2
      Contact( #qErrAcquiringTimeOut )
      I_Contact( #sResetFaults )
   END_RUNG wire#w4
   RUNG wire#w2
      Contact( #TriggerEnableTimeout.Q )
      wire#w5
      Coil( #qErrTriggerEnableTimeout )
   END_RUNG
   RUNG wire#w2
      Contact( #qErrTriggerEnableTimeout )
      I_Contact( #sResetFaults )
   END_RUNG wire#w5
   RUNG wire#w1
      Contact( #iStartJobSelection )
      Contact( #iInsightCamera_Input.iCommandFailed )
      wire#w6
      Coil( #qErrJobSelection )
   END_RUNG
   RUNG wire#w1
      Contact( #qErrJobSelection )
      I_Contact( #sResetFaults )
   END_RUNG wire#w6
   RUNG wire#w1
      Contact( #iStartInspection )
      Contact( #iStartJobSelection )
      wire#w7
      Coil( #qErrBothStartOn )
   END_RUNG
   RUNG wire#w1
      Contact( #qErrBothStartOn )
      I_Contact( #sResetFaults )
   END_RUNG wire#w7
   RUNG wire#w1
      Contact( #sPrgmNumTimer.Q )
      Contact( #iInsightCamera_Input.iSystemOnline )
      { S7_Templates := "SrcType := Int" } NE_Contact(in1 := #iJobID, in2 := #sVisionInputCmdControlIP)
      wire#w8
      Coil( #qErrJobIDEchoMismatch )
   END_RUNG
   RUNG wire#w1
      Contact( #qErrJobIDEchoMismatch )
      I_Contact( #sResetFaults )
   END_RUNG wire#w8
   RUNG wire#w1
      Contact( #sSetUserDataAckTimer.Q )
      wire#w9
      Coil( #qErrSetUserDataAckNtRcvd )
   END_RUNG
   RUNG wire#w1
      Contact( #qErrSetUserDataAckNtRcvd )
      I_Contact( #sResetFaults )
   END_RUNG wire#w9
   RUNG wire#w1
      Contact( #iStartInspection )
      { S7_Templates := "SrcType := Int" } NE_Contact(in1 := #iJobID, in2 := #iqRunningJobID)
      Coil( #qMsgJobIDMismatch )
   END_RUNG
   // the same network as SCL:
   #_w1 := true AND #iStartInspection;
   #qErrTriggerTimeOut := #_w1 AND (#TriggerTimeout.Q OR (#qErrTriggerTimeOut AND NOT #sResetFaults));
   #qErrAcquiringTimeOut := #_w1 AND (#AcquiringTimeOut.Q OR (#qErrAcquiringTimeOut AND NOT #sResetFaults));
   #qErrTriggerEnableTimeout := #_w1 AND (#TriggerEnableTimeout.Q OR (#qErrTriggerEnableTimeout AND NOT #sResetFaults));
   #qErrJobSelection := true AND ((#iStartJobSelection AND #iInsightCamera_Input.iCommandFailed) OR (#qErrJobSelection AND NOT #sResetFaults));
   #qErrBothStartOn := true AND ((#iStartInspection AND #iStartJobSelection) OR (#qErrBothStartOn AND NOT #sResetFaults));
   #qErrJobIDEchoMismatch := true AND ((#sPrgmNumTimer.Q AND #iInsightCamera_Input.iSystemOnline AND (#iJobID <> #sVisionInputCmdControlIP)) OR (#qErrJobIDEchoMismatch AND NOT #sResetFaults));
   #qErrSetUserDataAckNtRcvd := true AND (#sSetUserDataAckTimer.Q OR (#qErrSetUserDataAckNtRcvd AND NOT #sResetFaults));
   #qMsgJobIDMismatch := true AND #iStartInspection AND (#iJobID <> #iqRunningJobID);
END_REGION
END_FUNCTION_BLOCK

// folder: SM-Modules

FUNCTION "PR_WriteDataSlave" : Void   // FC19, LAD
TITLE = Write Data To Profinet Device
{ S7_Optimized_Access := 'TRUE' }
AUTHOR : GST
FAMILY : SM
NAME : SM0304022002
VERSION : 0.1
   VAR_INPUT
      iNumberOfBytes : Int;   // Number Of Bytes Configured In Hardware
      iSourceStruct : Variant;   // Source Data Structure
   END_VAR
   VAR_OUTPUT
      iOutputAddress : ANY;   // Output Data Address P#Q120.0 BYTE 71
   END_VAR
   VAR_TEMP
      tRetVal : Int;   // Ret Value
      tSrcMovBlck : Array[0..512] of Byte;   // Source Data ARRAY
      tPOS : DInt;   // POS
   END_VAR
BEGIN

REGION Network 1: Header
   // ==============================================================================
   //  Company: Precision Automation & Robotics India Ltd. 
   // ------------------------------------------------------------------------------
   //  Item Code: SM0304022002
   //  Author/Created by: GST
   //  Reviewed/Checked by: Atul P
   //  First Release on: 05-June-2018
   //  Latest update on: 
   // ------------------------------------------------------------------------------
   //  Tested with: CPU firmware, model or simulator testing
   //  Engineering/Editor: TIA Portal V15.1
   // ------------------------------------------------------------------------------
   //  Restrictions: 
   //  Dependencies/Requirements:
   //  This block uses following standard "Siemens" functions:
   // MOVE_BLK_VARIANT
   // Serialize
   // may lead to CPU going to STOP mode.
   // ------------------------------------------------------------------------------
   //  Change Log:
   //  Ver.	Date		Changed by		Details of changes
   //  1.0	05-June-2018	GST                               	First release version
   // ------------------------------------------------------------------------------
   //  Functionality:  This block is used for interface of Write Data From Structure Data To Profinet Device
   // 
   //  Inputs
   // iNumberOfBytes	Int
   // iSourceStruct	Variant
   // 
   //  Outputs
   // iOutputAddress	Any
   // 
   //  In-outs
   //  
   // ------------------------------------------------------------------------------
   //  Errors reported:
   //  1. 
   //  Messages reported:
   //  1. 
   // ==============================================================================
END_REGION

REGION Network 2: Serialize Structure Input Into Array
   // Serialize Structure Input Into Array
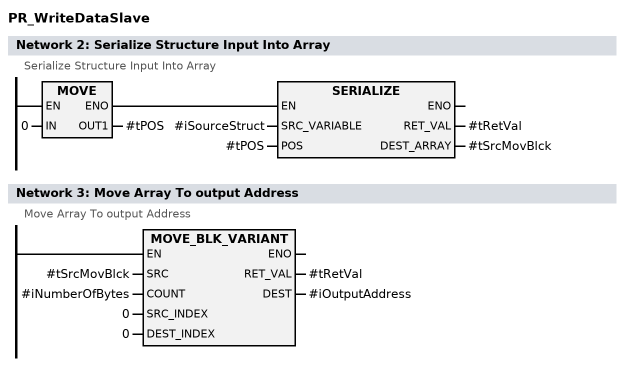
   // no SCL statement known for Serialize: written as a call
   #tPOS := 0;
   #tRetVal := Serialize(SRC_VARIABLE := #iSourceStruct, POS := #tPOS, DEST_ARRAY => #tSrcMovBlck);
END_REGION

REGION Network 3: Move Array To output Address
   // Move Array To output Address
   #tRetVal := MOVE_BLK_VARIANT(SRC := #tSrcMovBlck,
                           COUNT := #iNumberOfBytes,
                           SRC_INDEX := 0,
                           DEST_INDEX := 0,
                           DEST => #iOutputAddress);
END_REGION
END_FUNCTION

FUNCTION "PR_ReadDataSlave" : Void   // FC20, LAD
TITLE = Read Data From Profinet Device
{ S7_Optimized_Access := 'TRUE' }
AUTHOR : GST
FAMILY : SM
NAME : SM0314022001
VERSION : 0.1
// |BLOCK:Cognex Scanner Module
// Item Code : SMxxxxx
// Owner:Precision Automation & Robotics India Ltd.
// Author: GST
// Release Date:05-June-2018
// Version:0.1
// V0.1-Initial release
// |=============================================================================|
// Block Description: This block is used for interface of Read Data From Profinet Device And Store Into Structure DATA
// |=============================================================================|
// Errors:
// 
// =============================================================================|
// Dependency:
// This block uses following standard "Siemens" functions:
// MOVE_BLK_VARIANT
// Deserialize
// may lead to CPU going to STOP mode.
// |
   VAR_INPUT
      iInputAddress : ANY;   // Input Hardware Address P#I120.0 BYTE 77
      iNumberOfBytes : Int;   // Input Number Of Bytes
   END_VAR
   VAR_OUTPUT
      qDestStruct : Variant;   // Destination Data Structure
   END_VAR
   VAR_TEMP
      tRetVal : Int;   // Ret Value
      tDestMovBlck : Array[0..512] of Byte;   // Destination Data Array
      tPOS : DInt;   // POS
   END_VAR
BEGIN

REGION Network 1: Header
   // ==============================================================================
   //  Company: Precision Automation & Robotics India Ltd. 
   // ------------------------------------------------------------------------------
   //  Item Code: SM0314022001
   //  Author/Created by: GST
   //  Reviewed/Checked by: Atul P
   //  First Release on: 05-June-2018
   //  Latest update on:
   // ------------------------------------------------------------------------------
   //  Tested with: CPU firmware, model or simulator testing
   //  Engineering/Editor: TIA Portal V15.1
   // ------------------------------------------------------------------------------
   //  Restrictions: 
   //  Dependencies/Requirements:
   // This block uses following standard "Siemens" functions:
   // MOVE_BLK_VARIANT
   // Deserialize
   // may lead to CPU going to STOP mode.
   // ------------------------------------------------------------------------------
   //  Change Log:
   //  Ver.	Date		Changed by		Details of changes
   //  1.0	05-June-2018	GST                                   	First release version
   // ------------------------------------------------------------------------------
   //  Functionality: This block is used for interface of Read Data From Profinet Device And Store Into Structure DATA
   // 
   //  Inputs
   //  iInputAddress	Any
   // iNumberOfBytes	Int
   // 
   //  Outputs
   // qDestStruct	Variant
   // 
   //  In-outs
   //  
   // ------------------------------------------------------------------------------
   //  Errors reported:
   //  1.
   //  Messages reported:
   //  1. 
   // ==============================================================================
END_REGION

REGION Network 2: Move Input Address Data To Destination Array
   // Move Input Address Data To Destination Array
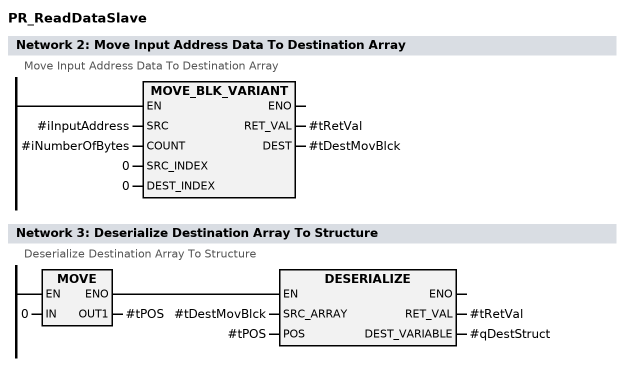
   #tRetVal := MOVE_BLK_VARIANT(SRC := #iInputAddress,
                           COUNT := #iNumberOfBytes,
                           SRC_INDEX := 0,
                           DEST_INDEX := 0,
                           DEST => #tDestMovBlck);
END_REGION

REGION Network 3: Deserialize Destination Array To Structure
   // Deserialize Destination Array To Structure
   // no SCL statement known for Deserialize: written as a call
   #tPOS := 0;
   #tRetVal := Deserialize(SRC_ARRAY := #tDestMovBlck, POS := #tPOS, DEST_VARIABLE => #qDestStruct);
END_REGION
END_FUNCTION